Fanuc KAREL source: KO00089.KL

PROGRAM KO00089
%NOLOCKGROUP
%ENVIRONMENT MIR
VAR
  P1: JOINTPOS
  P2: XYZWPREXT
  F: BOOLEAN
  OUT: POSITION
BEGIN
  F = TRUE
  OUT = MIRROR(P1, P2, F)
END KO00089
